(* IEC 61131-3 sources: rusty/tests/lit/single/parse_errors, 3 files *)

(* ---- error_format_none.st ---- *)
// RUN: not %COMPILE %s --error-format none 2>&1 | %CHECK %s
//
// With the error format none, parse errors are not printed. Only the abort line is printed.

FUNCTION foo : BOOL
VAR_INPUT
    in : BOOL;
    in2
END_VAR
;
END_FUNCTION

// CHECK-NOT: {{.+}}
// CHECK: error: Compilation aborted due to critical parse errors
// CHECK-NOT: {{.+}}

(* ---- reported_once_clang.st ---- *)
// RUN: not %COMPILE %s --error-format clang 2>&1 | %CHECK %s
//
// A parse error is reported once, in the clang format. The abort that follows does not repeat it.

FUNCTION foo : BOOL
VAR_INPUT
    in : BOOL;
    // CHECK: {{.*}}reported_once_clang.st:[[@LINE+1]]:{{[0-9]+}}:{{.*}}: error[E006]: Missing expected Token KeywordColon or KeywordComma
    in2
    // CHECK-NEXT: {{.*}}reported_once_clang.st:[[@LINE+4]]:1:{{.*}}: error[E006]: Missing expected Token KeywordColon
    // CHECK-NEXT: {{.*}}reported_once_clang.st:[[@LINE+3]]:1:{{.*}}: error[E007]: Unexpected token: expected DataTypeDefinition but found KeywordEndVar
    // CHECK-NEXT: {{.*}}reported_once_clang.st:[[@LINE+2]]:1:{{.*}}: error[E006]: Missing expected Token [KeywordSemicolon]
    // CHECK-NEXT: {{.*}}reported_once_clang.st:[[@LINE+1]]:1:{{.*}}: error[E007]: Unexpected token: expected KeywordSemicolon but found 'END_VAR'
END_VAR
;
END_FUNCTION

// CHECK-NEXT: error: Compilation aborted due to critical parse errors
// CHECK-NOT: {{.*}} at: {{.*}}

(* ---- reported_once_rich.st ---- *)
// RUN: not %COMPILE %s 2>&1 | %CHECK %s
//
// A parse error is reported once, in the rich format. The abort that follows does not repeat it
// in a "Details:" block. The rich reporter always writes color codes, so the error line allows them.

FUNCTION foo : BOOL
VAR_INPUT
    in : BOOL;
    in2
END_VAR
;
END_FUNCTION

// CHECK: {{.*}}error[E006]{{.*}}: Missing expected Token KeywordColon or KeywordComma{{.*}}
// CHECK: error: Compilation aborted due to critical parse errors.
// CHECK-NEXT: Hint: You can use `plc explain <ErrorCode>` for more information
